TYPE ST_MB_ReadRegs :
STRUCT
END_STRUCT
END_TYPE

(* stored: Version 1.1.0.1, ProductVersion 3.1.4024.13
   DUT ST_MB_ReadRegs: Id {ee3397d1-2360-4b44-84f6-8873fc2ec01e} *)
